(* CODESYS project candidate.project

Project tree, tasks and I/O mapping:
  CODESYS_Control_Win_x64 : CODESYS Control Win V3 x64, CODESYS, version 3.5.22.40
    application Application
      libraries: Standard, 3.5.22.0 (System)
      task MainTask (cyclic, interval t#50ms, priority 1) calls PLC_PRG
      program PLC_PRG [ST]
      function block FB_TemperatureControl [ST]
*)

// CODESYS_Control_Win_x64/Application/PLC_PRG
PROGRAM PLC_PRG
VAR
END_VAR

;

END_PROGRAM

// CODESYS_Control_Win_x64/Application/FB_TemperatureControl
FUNCTION_BLOCK FB_TemperatureControl

VAR_INPUT
    TemperatureSensorInput : REAL;
    SetTemperature : REAL;
END_VAR
VAR_OUTPUT
    CurrentTemperature : REAL;
    SetTempDisplay : REAL;
    HeaterStatus : BOOL;
    OverheatProtection : BOOL;
    HeaterOutput : BOOL;
END_VAR
VAR
    sensor_fault : BOOL;
    heater_request : BOOL;
    overheat_active : BOOL;
    tmp_heater_in : BOOL;
    HeatingTimer : TON;
    CoolingTimer : TON;
END_VAR

sensor_fault := (TemperatureSensorInput < 0.0) OR (TemperatureSensorInput > 100.0);
heater_request := (NOT sensor_fault) AND (TemperatureSensorInput < SetTemperature);


tmp_heater_in := heater_request AND NOT overheat_active;


HeatingTimer(IN := tmp_heater_in, PT := T#5S1MS);
IF HeatingTimer.Q THEN
    overheat_active := TRUE;
    tmp_heater_in := FALSE;
END_IF;


CoolingTimer(IN := overheat_active, PT := T#3S);
IF overheat_active AND CoolingTimer.Q THEN
    overheat_active := FALSE;
END_IF;

HeaterOutput := heater_request AND NOT overheat_active;


IF HeaterOutput AND NOT tmp_heater_in THEN
    HeatingTimer(IN := TRUE, PT := T#5S1MS);
ELSIF (NOT HeaterOutput) AND tmp_heater_in THEN
    HeatingTimer(IN := FALSE, PT := T#5S1MS);
END_IF;

CurrentTemperature := TemperatureSensorInput;
SetTempDisplay := SetTemperature;
HeaterStatus := HeaterOutput;
OverheatProtection := overheat_active;

END_FUNCTION_BLOCK
